(* PLC project Simulatie Sorteer Station, CODESYS CODESYS V3.5 SP16 Patch 7, author Rene Potters/Gerard Harkema *)
(* stored: creationDateTime 2026-11-25T11:59:04.5501741, version 0.1.0, modificationDateTime 2026-11-25T11:44:06.263536, organization Avans *)
(* Simulatie voor opstelling Sorteer Station. *)

VAR_GLOBAL  (* GVL *)
  Ix_Resetknop : BOOL;  (* Indrukken resetknop *)
  Ix_Hand : BOOL;  (* Keuzeknop staat op hand *)
  Ix_Auto : BOOL;  (* Keuzeknop staat op auto *)
  Ix_Noodstop : BOOL;  (* Indrukken noodstop *)
  Ix_MagazijnLeeg : BOOL;  (* Bekers magazijn zijn op *)
  Ix_UitstoterBekerIn : BOOL;  (* Beker is uit dekselmagazijn gestoten *)
  Ix_UitstoterBekerUit : BOOL;  (* Uitstoter Beker haalt nieuwe beker op *)
  Ix_Stopknop : BOOL := TRUE;  (* Indrukken startknop *)
  Ix_Startknop : BOOL;  (* Indrukken stopknop *)
  Ix_PersluchtAanwezig : BOOL;  (* Perslucht is aanwezig *)
  Ix_VacuumAanwezig : BOOL;  (* Werkstuk door overzetter opgepakt *)
  Ix_OverzetterIsLinks : BOOL;  (* Overzetter haalt beker op(linker pos.) *)
  Ix_OverzetterIsRechts : BOOL;  (* Overzetter plaatst beker op sorteerpositie *)
  Ix_BekerAanwezig : BOOL;  (* Beker aanwezig op detectiepositie *)
  Ix_BekerMetaal : BOOL;  (* Beker is van aluminium *)
  Ix_BekerReflecteerd : BOOL;  (* Beker reflecteert en is dus niet zwart *)
  Ix_BekerInGoot : BOOL;  (* Product is naar een van de goten gegaan *)
  Ix_UitvoerGoot1IsIn : BOOL;  (* Pusher uitvoergoot 1 is in *)
  Ix_UitvoerGoot2IsIn : BOOL;  (* Pusher uitvoergoot 2 is in *)
  Ix_StationAfvoerVrij : BOOL;  (* Beker afvoeren is bezig *)
  Ix_UitvoerGoot1IsUit : BOOL;  (* Pusher uitvoergoot 1 is uit *)
  Ix_UitvoerGoot2IsUit : BOOL;  (* Pusher uitvoergoot 2 is uit *)
  Qx_BekerUitstoten : BOOL;  (* Beker uit magazijn stoten *)
  Qx_VacuumAan : BOOL;  (* Beker oppakken *)
  Qx_BekerLossen : BOOL;  (* Beker loslaten *)
  Qx_OverzetterLinks : BOOL;  (* Overzetter naar bekermagazijn *)
  Qx_OverzetterRechts : BOOL;  (* Overzetter naar sorteerpositie *)
  Qx_MotorAfvoerAan : BOOL;  (* Transportband aan *)
  Qx_UitvoerGoot1Uit : BOOL;  (* Pusher goot 1 uit *)
  Qx_UitvoerGoot2Uit : BOOL;  (* Pusher goot 2 uit *)
  Qx_StopperUit : BOOL;  (* Beker stoppen op band voor detectie *)
  Qx_StationBezet : BOOL;  (* Uitsorteren is bezet *)
  Qx_GeleLamp : BOOL;  (* Visualisatie invisible Gele vlak *)
  Qx_GroeneLamp : BOOL;  (* Visualisatie invisible groene vlak *)
  Qx_RodeLamp : BOOL;  (* Visualisatie invisible rode vlak *)
END_VAR

CONFIGURATION Device
  RESOURCE ApplicationLadder ON PLC
    TASK MainTask(INTERVAL := T#20ms, PRIORITY := 1);
    TASK Simulatie(INTERVAL := T#50ms, PRIORITY := 1);
    PROGRAM BedieningPrg WITH MainTask : BedieningPrg;
    PROGRAM HoofdPrg WITH MainTask : HoofdPrg;
    PROGRAM MagazijnPrg WITH MainTask : MagazijnPrg;
    PROGRAM OverzetterPrg WITH MainTask : OverzetterPrg;
    PROGRAM SorterenPrg WITH MainTask : SorterenPrg;
    PROGRAM SignaleringPrg WITH MainTask : SignaleringPrg;
    PROGRAM MagazijnSim WITH Simulatie : MagazijnSim;
    PROGRAM OverzetterSim WITH Simulatie : OverzetterSim;
    PROGRAM SorterenSim WITH Simulatie : SorterenSim;
  END_RESOURCE
  RESOURCE ApplicationSt ON PLC
    TASK MainTask(INTERVAL := T#20ms, PRIORITY := 1);
    TASK Simulatie(INTERVAL := T#20ms, PRIORITY := 1);
    PROGRAM Main WITH MainTask : Main;
    PROGRAM MagazijnSim WITH Simulatie : MagazijnSim;
    PROGRAM OverzetterSim WITH Simulatie : OverzetterSim;
    PROGRAM SorterenSim WITH Simulatie : SorterenSim;
  END_RESOURCE
  RESOURCE MagazijnTest ON PLC
    TASK MainTask(INTERVAL := T#20ms, PRIORITY := 1);
    TASK Simulatie(INTERVAL := T#20ms, PRIORITY := 1);
    PROGRAM MagazijnTest WITH MainTask : MagazijnTest;
    PROGRAM MagazijnSim WITH Simulatie : MagazijnSim;
  END_RESOURCE
  RESOURCE OverzetterTest ON PLC
    TASK MainTask(INTERVAL := T#20ms, PRIORITY := 1);
    TASK Simulatie(INTERVAL := T#20ms, PRIORITY := 1);
    PROGRAM OverzetterTest WITH MainTask : OverzetterTest;
    PROGRAM OverzetterSim WITH Simulatie : OverzetterSim;
  END_RESOURCE
  RESOURCE SorteerTest ON PLC
    TASK MainTask(INTERVAL := T#20ms, PRIORITY := 1);
    TASK Simulatie(INTERVAL := T#20ms, PRIORITY := 1);
    PROGRAM SorteerTest WITH MainTask : SorteerTest;
    PROGRAM SorterenSim WITH Simulatie : SorterenSim;
  END_RESOURCE
  RESOURCE UitvoerGootTest ON PLC
    TASK MainTask(INTERVAL := T#20ms, PRIORITY := 1);
    TASK Simulatie(INTERVAL := T#20ms, PRIORITY := 1);
    PROGRAM UitvoerGootTest WITH MainTask : UitvoerGootTest;
    PROGRAM SorterenSim WITH Simulatie : SorterenSim;
  END_RESOURCE
END_CONFIGURATION

CONFIGURATION Basic
END_CONFIGURATION

CONFIGURATION <Empty>
END_CONFIGURATION

CONFIGURATION <Empty>
END_CONFIGURATION

CONFIGURATION <Empty>
END_CONFIGURATION

CONFIGURATION <Empty>
END_CONFIGURATION

CONFIGURATION <Empty>
END_CONFIGURATION

CONFIGURATION <Empty>
END_CONFIGURATION

CONFIGURATION <Empty>
END_CONFIGURATION

CONFIGURATION <Empty>
END_CONFIGURATION

CONFIGURATION <Empty>
END_CONFIGURATION

CONFIGURATION <Empty>
END_CONFIGURATION

CONFIGURATION <Empty>
END_CONFIGURATION
